Fanuc KAREL source: kb00068.compact.KL

PROGRAM KB00068
%STACKSIZE=65535
%PRIORITY=65535
%NOLOCKGROUP
%ENVIRONMENT FDEV
VAR
P1 : STRING[80]
P2 : INTEGER
BEGIN
P1='A'
P2=1
DISMOUNT_DEV(P1,P2)
END KB00068
